Universal Robots URScript: PrecProg.script

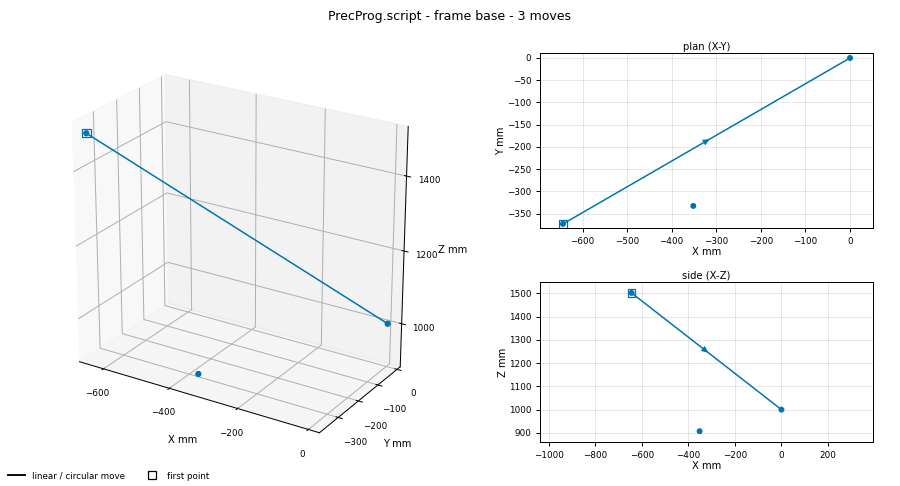
[picture p0: tool path of PrecProg.script in frame base, 3 of 6 moves have a stored position in this frame; points joined in program order, loops and branches not executed]
def PrecProg():
  # Global parameters:
  global speed_ms    = 0.250
  global speed_rads  = 0.750
  global accel_mss   = 1.200
  global accel_radss = 1.200
  global blend_radius_m = 0.000

  #--------------------------
  # Add any default subprograms here
  # For example, to drive a gripper as a program call:
  # def Gripper_Open():
  #   ...
  # end
  #
  # Example to drive a spray gun:
  def SprayOn(value):
    # use the value as an output:
    DO_SPRAY = 5
    if value == 0:
      set_standard_digital_out(DO_SPRAY, False)
    else:
      set_standard_digital_out(DO_SPRAY, True)
    end
  end

  # Example to synchronize 2
  def Synchronize():
    # Use the following digital output to signal the state of the robot:
    DO_SYNC = 1

    # Use the following digital input to get the state of another robot:
    DI_SYNC = 1

    if (get_standard_digital_out(DO_SYNC) == get_standard_digital_in(DI_SYNC)):
      set_standard_digital_out(DO_SYNC, not (get_standard_digital_out(DI_SYNC)))
      sleep(0.1)
      thread Thread_wait_1():
        while (True):
          sleep(0.01)
        end
      end
      if (get_standard_digital_out(DO_SYNC) != get_standard_digital_in(DI_SYNC)):
        global thread_handler_1=run Thread_wait_1()
        while (get_standard_digital_out(DO_SYNC) != get_standard_digital_in(DI_SYNC)):
          sync()
        end
        kill thread_handler_1
      end
    else:
      if (get_standard_digital_out(DO_SYNC) != get_standard_digital_in(DI_SYNC)):
        set_standard_digital_out(DO_SYNC, not (get_standard_digital_out(DO_SYNC)))
      end
    end
  end

  #
  # Example to move an external axis
  def MoveAxis(value):
    # use the value as an output:
    DO_AXIS_1 = 1
    DI_AXIS_1 = 1
    if value <= 0:
      set_standard_digital_out(DO_AXIS_1, False)

      # Wait for digital input to change state
      #while (get_standard_digital_in(DI_AXIS_1) != False):
      #  sync()
      #end
    else:
      set_standard_digital_out(DO_AXIS_1, True)

      # Wait for digital input to change state
      #while (get_standard_digital_in(DI_AXIS_1) != True):
      #  sync()
      #end
    end
  end
  #--------------------------


  # Main program:
  # Program generated by RoboDK v6.0.7 for ABB IRB 120-3/0.6 on XX/XX/XXXX 18:00:00
  # Using nominal kinematics.
  # Using Ref. Frame P: p[0.000000, -0.000001, 1.000000, 1.570792, -0.005162, 0.008546]
  # set_reference(p[0.000000, -0.000001, 1.000000, 1.570792, -0.005162, 0.008546])
  # Using TCP Tool P: p[0.000125, -0.000375, 0.123457, -0.789761, -0.000001, 0.000002]
  set_tcp(p[0.000125, -0.000375, 0.123457, -0.789761, -0.000001, 0.000002])
  movej([0.215471, -0.797247, 1.377087, -0.008727, 0.008726, 3.141593],1.20000,0.75000,0,0.0000)
  movel(p[-0.644182, -0.372923, 1.501372, 1.397179, 2.288562, 1.360920],accel_mss,speed_ms,0,0.000)
  movel(p[0.000505, -0.000250, 0.999504, -1.570776, -0.008546, -0.005299],accel_mss,speed_ms,0,0.000)
  movej([-0.215468, 0.797240, -1.377065, 0.008727, -0.000002, -3.141593],1.20000,0.75000,0,0.0000)
  movej([-0.215468, 0.797240, -1.377065, 0.008727, -0.000002, -3.141593],1.20000,0.75000,0,0.0000)
  speed_ms    = 0.0667
  sleep(0.002)
  sleep(1.000)
  movel(p[-0.351510, -0.332461, 0.906789, 0.761248, 2.011888, 1.655391],accel_mss,speed_ms,0,0.000)
  # End of main program
end

PrecProg()
